// TIA Portal V20 export
// export: Created 2026-10-12T05:14:46.445642Z, ExportSetting WithDefaults, DisplayName Totally Integrated Automation Portal, DisplayVersion V20, DisplayName TIA Portal Openness, DisplayVersion V20, DisplayName TIA Portal Teamcenter Gateway, DisplayVersion V20, DisplayName TIA Portal Version Control Interface, DisplayVersion V20, DisplayName SINAMICS Startdrive Advanced, DisplayVersion V20 SP1 Update 2, DisplayName SINAMICS Startdrive G110M, G120, G120C, G120D, G120P, G115D, DisplayVersion V20 SP1 Update 2, DisplayName SINAMICS Startdrive G130, G150, S120, S150, SINAMICS MV, G220, S200, S210, DisplayVersion V20 SP1 Update 2, DisplayName STEP 7 Professional, DisplayVersion V20, DisplayName STEP 7 Safety, DisplayVersion V20, DisplayName WinCC Basic/Comfort/Advanced, DisplayVersion V20, DisplayName WinCC Professional, DisplayVersion V20, DisplayName WinCC Unified, DisplayVersion V20
FUNCTION "FRK_JsonReadRecord" : Bool   // FC122, SCL
{ S7_Optimized_Access := 'TRUE' }
VERSION : 0.1
// stored: AutoNumber true, IsIECCheckEnabled false, SetENOAutomatically false, UDAEnableTagReadback false
   VAR_INPUT
      Count : Int;
      Fields : Array[1..9] of "FRK_JsonField";
   END_VAR
   VAR_IN_OUT
      Data : "ST_ConfigRecord";
   END_VAR
   VAR_TEMP
      Candidate : "ST_ConfigRecord";
      Index : Int;
      Found : Int;
      Ok : Bool;
   END_VAR
BEGIN

   #FRK_JsonReadRecord := FALSE;
   IF #Count <> 6 THEN
       RETURN;
   END_IF;
   #Found := 0;
   FOR #Index := 1 TO #Count DO
       IF #Fields[#Index].Key = 'scope' THEN
           #Found := #Index;
       END_IF;
   END_FOR;
   IF #Found = 0 THEN
       RETURN;
   END_IF;
   IF #Fields[#Found].Quoted <> TRUE THEN
       RETURN;
   END_IF;
   IF LEN(#Fields[#Found].Text) > 80 OR STRING_TO_WSTRING(WSTRING_TO_STRING(#Fields[#Found].Text)) <> #Fields[#Found].Text THEN
       RETURN;
   END_IF;
   #Candidate.Scope := WSTRING_TO_STRING(#Fields[#Found].Text);
   #Found := 0;
   FOR #Index := 1 TO #Count DO
       IF #Fields[#Index].Key = 'key' THEN
           #Found := #Index;
       END_IF;
   END_FOR;
   IF #Found = 0 THEN
       RETURN;
   END_IF;
   IF #Fields[#Found].Quoted <> TRUE THEN
       RETURN;
   END_IF;
   IF LEN(#Fields[#Found].Text) > 160 OR STRING_TO_WSTRING(WSTRING_TO_STRING(#Fields[#Found].Text)) <> #Fields[#Found].Text THEN
       RETURN;
   END_IF;
   #Candidate.WriteKey := WSTRING_TO_STRING(#Fields[#Found].Text);
   #Found := 0;
   FOR #Index := 1 TO #Count DO
       IF #Fields[#Index].Key = 'rev' THEN
           #Found := #Index;
       END_IF;
   END_FOR;
   IF #Found = 0 THEN
       RETURN;
   END_IF;
   IF #Fields[#Found].Quoted <> FALSE THEN
       RETURN;
   END_IF;
   #Ok := "FRK_ConfigDecode"(Text := #Fields[#Found].Text, Storage := 4, Minimum := 0.0, Maximum := 4294967295.0, MaxLength := 0, Value := "FRK_ConfigScratch".Value);
   IF NOT #Ok THEN
       RETURN;
   END_IF;
   #Candidate.Revision := LINT_TO_UDINT("FRK_ConfigScratch".Value.Number);
   #Found := 0;
   FOR #Index := 1 TO #Count DO
       IF #Fields[#Index].Key = 'kind' THEN
           #Found := #Index;
       END_IF;
   END_FOR;
   IF #Found = 0 THEN
       RETURN;
   END_IF;
   IF #Fields[#Found].Quoted <> FALSE THEN
       RETURN;
   END_IF;
   #Ok := "FRK_ConfigDecode"(Text := #Fields[#Found].Text, Storage := 4, Minimum := 0.0, Maximum := 1.0, MaxLength := 0, Value := "FRK_ConfigScratch".Value);
   IF NOT #Ok THEN
       RETURN;
   END_IF;
   #Candidate.Kind := LINT_TO_DINT("FRK_ConfigScratch".Value.Number);
   #Found := 0;
   FOR #Index := 1 TO #Count DO
       IF #Fields[#Index].Key = 'type' THEN
           #Found := #Index;
       END_IF;
   END_FOR;
   IF #Found = 0 THEN
       RETURN;
   END_IF;
   IF #Fields[#Found].Quoted <> FALSE THEN
       RETURN;
   END_IF;
   #Ok := "FRK_ConfigDecode"(Text := #Fields[#Found].Text, Storage := 4, Minimum := 0.0, Maximum := 3.0, MaxLength := 0, Value := "FRK_ConfigScratch".Value);
   IF NOT #Ok THEN
       RETURN;
   END_IF;
   #Candidate.ValueType := LINT_TO_DINT("FRK_ConfigScratch".Value.Number);
   #Found := 0;
   FOR #Index := 1 TO #Count DO
       IF #Fields[#Index].Key = 'value' THEN
           #Found := #Index;
       END_IF;
   END_FOR;
   IF #Found = 0 THEN
       RETURN;
   END_IF;
   IF #Fields[#Found].Quoted <> TRUE THEN
       RETURN;
   END_IF;
   IF LEN(#Fields[#Found].Text) > 80 OR STRING_TO_WSTRING(WSTRING_TO_STRING(#Fields[#Found].Text)) <> #Fields[#Found].Text THEN
       RETURN;
   END_IF;
   #Candidate.ValueText := WSTRING_TO_STRING(#Fields[#Found].Text);
   #Data := #Candidate;
   #FRK_JsonReadRecord := TRUE;
END_FUNCTION
